# EPICS autosave request: iocBoot/iocUSBTEMP-AI/auto_settings.req
file "USBTEMP_AI_settings.req", P=$(P)
